Universal Robots URScript: MAIN_1.script

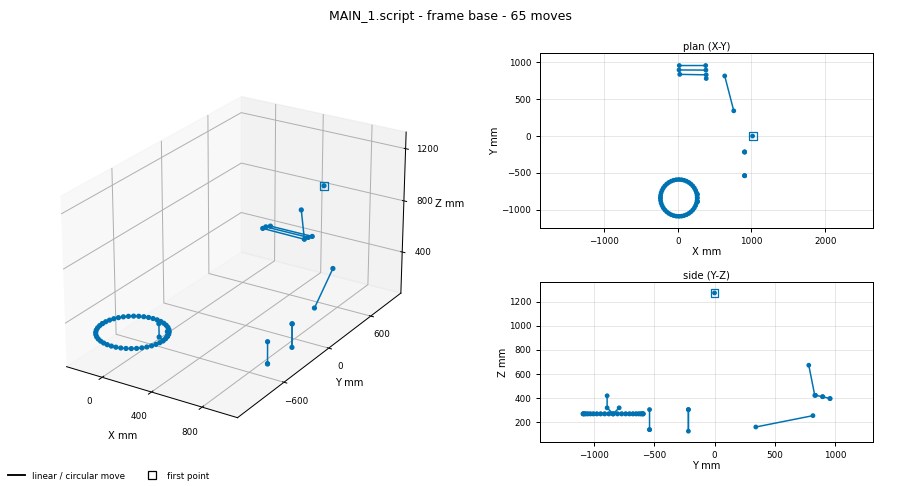
[picture p0: tool path of MAIN_1.script in frame base, 65 of 76 moves have a stored position in this frame; points joined in program order, loops and branches not executed]
def MAIN_1():
  # Global parameters:
  global speed_ms    = 0.300
  global speed_rads  = 0.750
  global accel_mss   = 3.000
  global accel_radss = 1.200
  global blend_radius_m = 0.001

  #--------------------------
  # Add any default subprograms here
  # For example, to drive a gripper as a program call:
  # def Gripper_Open():
  #   ...
  # end
  #
  # Example to drive a spray gun:
  def SprayOn(value):
    # use the value as an output:
    DO_SPRAY = 5
    if value == 0:
      set_standard_digital_out(DO_SPRAY, False)
    else:
      set_standard_digital_out(DO_SPRAY, True)
    end
  end

  # Example to drive an extruder:
  def Extruder(value):
    # use the value as an output:
    if value < 0:
      # stop extruder
    else:
      # start extruder
    end
  end

  # Example to move an external axis
  def MoveAxis(value):
    # use the value as an output:
    DO_AXIS_1 = 1
    DI_AXIS_1 = 1
    if value <= 0:
      set_standard_digital_out(DO_AXIS_1, False)

      # Wait for digital input to change state
      #while (get_standard_digital_in(DI_AXIS_1) != False):
      #  sync()
      #end
    else:
      set_standard_digital_out(DO_AXIS_1, True)

      # Wait for digital input to change state
      #while (get_standard_digital_in(DI_AXIS_1) != True):
      #  sync()
      #end
    end
  end
  #--------------------------

  # Subprogram PROG1_withaverylongnameandspecialcharacters
  def PROG1_withaverylongnameandspecialcharacters():
    # This is a subprogram call to PROG_1
    # set_reference(p[0.000000, 1.000000, 0.000000, 0.000000, 0.000000, 0.000000])
    set_tcp(p[0.000000, 0.000000, 0.200000, 0.000000, 0.000000, 0.000000])
    movej([-0.000000, 0.000000, 0.000000, 0.000000, 0.000000, -0.000000],accel_radss,speed_rads,0,blend_radius_m)
  end


  # Main program:
  # Program generated by RoboDK v5.6.9 for RoboDK Industrial on 26/02/2024 09:58:20
  # Using nominal kinematics.
  movej([-0.000000, 0.000000, 0.000000, 0.000000, 0.000000, -0.000000],accel_radss,speed_rads,0,0)
  movej([0.000000, 0.056047, -0.269194, 0.000000, 0.213148, -0.000000],accel_radss,speed_rads,0,0)
  movel(p[1.015000, 0.000000, 1.272000, 0.000000, 1.570796, 0.000000],accel_mss,speed_ms,0,blend_radius_m)
  set_standard_digital_out(5, True)
  set_standard_digital_out(5, True)
  set_standard_digital_out(5, 0.5)
  set_standard_digital_out(5, true)
  set_standard_digital_out(5, True)
  set_standard_digital_out(5, True)
  set_standard_digital_out(5, 0.5)
  set_standard_digital_out(5, true)
  var = val
  var = val
  while (get_standard_digital_in(5) != True):
    sync()
  end
  while (get_standard_digital_in(5) != True):
    sync()
  end
  while (get_standard_digital_in(5) != 0.5):
    sync()
  end
  while (get_standard_digital_in(5) != true):
    sync()
  end
  while (get_standard_digital_in(5) != True):
    sync()
  end
  while (var != val):
    sync()
  end
  while (var != val):
    sync()
  end
  popup("Message","Message",False,False,blocking=True)
  REMOTE_PROG_CALL_171()
  # CODE_INSERT_172
  # Insert Comment
  # set_reference(p[0.719013, -0.664003, 0.000000, 0.000000, 0.000000, 0.000000])
  set_tcp(p[0.129073, 0.000000, 0.085477, 0.000000, 0.398790, 0.000000])
  accel_radss = 13.963
  speed_rads  = 8.727
  blend_radius_m = 0.010
  movej([-0.511943, 0.814667, -0.000428, 0.463308, 0.443239, -0.901183],accel_radss,speed_rads,0,blend_radius_m)
  blend_radius_m = 0.000
  accel_mss   = 0.200
  speed_ms    = 0.100
  movel(p[0.906799, -0.538504, 0.139112, -0.000082, 3.138451, 0.000110],accel_mss,speed_ms,0,blend_radius_m)
  set_standard_digital_out(5, True)
  PICK_PART_111()
  blend_radius_m = 0.010
  accel_mss   = 0.600
  speed_ms    = 0.300
  movel([-0.511943, 0.814667, -0.000427, 0.463312, 0.443239, -0.901187],accel_mss,speed_ms,0,0)
  movel(p[0.906285, -0.216481, 0.305347, 0.000027, 3.138364, -0.000055],accel_mss,speed_ms,0,blend_radius_m)
  blend_radius_m = 0.000
  accel_mss   = 0.200
  speed_ms    = 0.100
  # MoveSearch command not implemented
  movel(p[0.906864, -0.216486, 0.126235, 0.000027, 3.138364, -0.000055],accel_mss,speed_ms,0,blend_radius_m)
  set_standard_digital_out(5, False)
  PLACE_PART_112()
  blend_radius_m = 0.010
  movel(p[0.906285, -0.216481, 0.305347, 0.000027, 3.138364, -0.000055],accel_mss,speed_ms,0,blend_radius_m)
  # set_reference(p[0.577670, 0.392250, 0.000000, 0.000000, 0.000000, 0.679972])
  blend_radius_m = 0.025
  accel_radss = 13.963
  speed_rads  = 8.727
  accel_mss   = 0.200
  speed_ms    = 0.100
  movej([0.910818, 0.797193, 0.120777, 1.164732, 0.347884, -1.618444],accel_radss,speed_rads,0,blend_radius_m)
  movec(p[0.884547, 0.696689, 0.231503, -2.018719, 2.221778, 0.218496],p[0.759304, 0.342075, 0.161073, -2.018719, 2.221778, 0.218496],accel_mss,speed_ms,blend_radius_m)
  # Circular movement using joint targets is not supported. Change the target type to cartesian or use a joint movement.
  blend_radius_m = 0.000
  accel_mss   = 0.200
  speed_ms    = 0.100
  movel(p[0.636704, 0.815780, 0.255156, -2.018719, 2.221778, 0.218496],accel_mss,speed_ms,0,blend_radius_m)
  movej([-0.000000, 0.000000, 0.000000, 0.000000, 0.000000, -0.000000],accel_radss,speed_rads,0,0)
  # set_reference(p[0.000000, 0.782714, 0.377610, 0.000000, 0.000000, 0.000000])
  movej([1.547688, 0.516645, -0.112204, -0.034631, 0.863575, 0.079372],accel_radss,speed_rads,0,0)
  movel(p[0.019898, 0.957021, 0.396618, 2.079600, -2.265750, 0.107759],accel_mss,speed_ms,0,blend_radius_m)
  movel(p[0.378402, 0.957130, 0.396607, 2.079600, -2.265750, 0.107759],accel_mss,speed_ms,0,blend_radius_m)
  movel(p[0.380996, 0.895077, 0.412492, 1.963520, -2.143933, 0.343573],accel_mss,speed_ms,0,blend_radius_m)
  movel(p[0.016551, 0.897073, 0.411836, 1.963520, -2.143933, 0.343573],accel_mss,speed_ms,0,blend_radius_m)
  movel(p[0.026434, 0.837238, 0.423682, -2.078092, 2.285598, 0.087159],accel_mss,speed_ms,0,blend_radius_m)
  movel(p[0.385448, 0.830764, 0.422747, -2.018705, 2.221797, 0.218488],accel_mss,speed_ms,0,blend_radius_m)
  movel(p[0.385448, 0.781089, 0.672861, -2.018705, 2.221797, 0.218488],accel_mss,speed_ms,0,blend_radius_m)
  movej([-0.000000, 0.000000, 0.000000, 0.000000, 0.000000, -0.000000],accel_radss,speed_rads,0,0)
  EVENT_PROG_START_101()
  blend_radius_m = 0.001
  speed_ms    = 1.000
  # set_reference(p[0.013637, -0.840080, 0.000000, 0.000000, 0.000000, -1.570796])
  # Show Tool 1
  movej([-1.188400, 0.422403, 0.467495, 0.666950, 0.631839, -1.724322],accel_radss,speed_rads,0,0)
  EVENT_PATH_APPROACH_102()
  movel(p[0.266896, -0.790185, 0.319999, 0.000002, 3.135432, -0.000684],accel_mss,speed_ms,0,blend_radius_m)
  movel(p[0.263637, -0.840080, 0.270000, 0.000002, 3.135432, -0.000684],accel_mss,speed_ms,0,blend_radius_m)
  EVENT_PATH_START_103()
  speed_ms    = 0.050
  movel(p[0.261092, -0.875659, 0.270000, 0.000006, 3.135571, -0.002052],accel_mss,speed_ms,0,blend_radius_m)
  movel(p[0.253510, -0.910513, 0.270000, -0.000018, 3.135814, -0.003393],accel_mss,speed_ms,0,blend_radius_m)
  movel(p[0.241045, -0.943934, 0.270000, -0.000015, 3.136179, -0.004625],accel_mss,speed_ms,0,blend_radius_m)
  movel(p[0.223950, -0.975240, 0.270000, -0.000013, 3.136648, -0.005803],accel_mss,speed_ms,0,blend_radius_m)
  movel(p[0.202574, -1.003795, 0.270000, -0.000012, 3.137222, -0.006844],accel_mss,speed_ms,0,blend_radius_m)
  movel(p[0.177352, -1.029017, 0.270000, -0.000013, 3.137883, -0.007749],accel_mss,speed_ms,0,blend_radius_m)
  movel(p[0.148797, -1.050393, 0.270000, -0.000015, 3.138614, -0.008518],accel_mss,speed_ms,0,blend_radius_m)
  movel(p[0.117491, -1.067488, 0.270000, -0.000018, 3.139415, -0.009096],accel_mss,speed_ms,0,blend_radius_m)
  movel(p[0.084070, -1.079953, 0.270000, 0.000006, 3.140269, -0.009482],accel_mss,speed_ms,0,blend_radius_m)
  movel(p[0.049216, -1.087535, 0.270000, 0.000002, 3.141141, -0.009676],accel_mss,speed_ms,0,blend_radius_m)
  movel(p[0.013637, -1.090080, 0.270000, 0.000002, -3.141141, 0.009676],accel_mss,speed_ms,0,blend_radius_m)
  movel(p[-0.021942, -1.087535, 0.270000, 0.000006, -3.140269, 0.009482],accel_mss,speed_ms,0,blend_radius_m)
  movel(p[-0.056796, -1.079953, 0.270000, -0.000018, -3.139415, 0.009096],accel_mss,speed_ms,0,blend_radius_m)
  movel(p[-0.090217, -1.067488, 0.270000, -0.000015, -3.138614, 0.008518],accel_mss,speed_ms,0,blend_radius_m)
  movel(p[-0.121523, -1.050393, 0.270000, -0.000013, -3.137883, 0.007749],accel_mss,speed_ms,0,blend_radius_m)
  movel(p[-0.150078, -1.029017, 0.270000, -0.000012, -3.137222, 0.006844],accel_mss,speed_ms,0,blend_radius_m)
  movel(p[-0.175300, -1.003795, 0.270000, -0.000013, -3.136648, 0.005803],accel_mss,speed_ms,0,blend_radius_m)
  movel(p[-0.196676, -0.975240, 0.270000, -0.000015, -3.136161, 0.004653],accel_mss,speed_ms,0,blend_radius_m)
  movel(p[-0.213771, -0.943934, 0.270000, -0.000018, -3.135796, 0.003393],accel_mss,speed_ms,0,blend_radius_m)
  movel(p[-0.226236, -0.910513, 0.270000, 0.000006, -3.135553, 0.002052],accel_mss,speed_ms,0,blend_radius_m)
  movel(p[-0.233818, -0.875659, 0.270000, 0.000002, -3.135432, 0.000684],accel_mss,speed_ms,0,blend_radius_m)
  movel(p[-0.236363, -0.840080, 0.270000, 0.000002, -3.135432, 0.000684],accel_mss,speed_ms,0,blend_radius_m)
  movel(p[-0.236363, -0.840080, 0.270000, -0.000002, -3.135432, -0.000684],accel_mss,speed_ms,0,0.000)
  movel(p[-0.233818, -0.804501, 0.270000, -0.000006, -3.135553, -0.002052],accel_mss,speed_ms,0,blend_radius_m)
  movel(p[-0.226236, -0.769647, 0.270000, 0.000018, -3.135814, -0.003393],accel_mss,speed_ms,0,blend_radius_m)
  movel(p[-0.213771, -0.736226, 0.270000, 0.000015, -3.136179, -0.004625],accel_mss,speed_ms,0,blend_radius_m)
  movel(p[-0.196676, -0.704920, 0.270000, 0.000013, -3.136648, -0.005803],accel_mss,speed_ms,0,blend_radius_m)
  movel(p[-0.175300, -0.676365, 0.270000, 0.000012, -3.137222, -0.006844],accel_mss,speed_ms,0,blend_radius_m)
  movel(p[-0.150078, -0.651143, 0.270000, 0.000013, -3.137883, -0.007749],accel_mss,speed_ms,0,blend_radius_m)
  movel(p[-0.121523, -0.629767, 0.270000, 0.000015, -3.138632, -0.008491],accel_mss,speed_ms,0,blend_radius_m)
  movel(p[-0.090217, -0.612672, 0.270000, 0.000018, -3.139433, -0.009068],accel_mss,speed_ms,0,blend_radius_m)
  movel(p[-0.056796, -0.600207, 0.270000, -0.000006, -3.140269, -0.009482],accel_mss,speed_ms,0,blend_radius_m)
  movel(p[-0.021942, -0.592625, 0.270000, -0.000002, -3.141141, -0.009676],accel_mss,speed_ms,0,blend_radius_m)
  movel(p[0.013637, -0.590080, 0.270000, -0.000002, 3.141141, 0.009676],accel_mss,speed_ms,0,blend_radius_m)
  movel(p[0.049216, -0.592625, 0.270000, -0.000006, 3.140269, 0.009454],accel_mss,speed_ms,0,blend_radius_m)
  movel(p[0.084070, -0.600207, 0.270000, 0.000018, 3.139433, 0.009068],accel_mss,speed_ms,0,blend_radius_m)
  movel(p[0.117491, -0.612672, 0.270000, 0.000015, 3.138614, 0.008518],accel_mss,speed_ms,0,blend_radius_m)
  movel(p[0.148797, -0.629767, 0.270000, 0.000013, 3.137883, 0.007749],accel_mss,speed_ms,0,blend_radius_m)
  movel(p[0.177352, -0.651143, 0.270000, 0.000012, 3.137222, 0.006844],accel_mss,speed_ms,0,blend_radius_m)
  movel(p[0.202574, -0.676365, 0.270000, 0.000013, 3.136648, 0.005803],accel_mss,speed_ms,0,blend_radius_m)
  movel(p[0.223950, -0.704920, 0.270000, 0.000015, 3.136179, 0.004625],accel_mss,speed_ms,0,blend_radius_m)
  movel(p[0.241045, -0.736226, 0.270000, 0.000018, 3.135796, 0.003393],accel_mss,speed_ms,0,blend_radius_m)
  movel(p[0.253510, -0.769647, 0.270000, -0.000006, 3.135553, 0.002052],accel_mss,speed_ms,0,blend_radius_m)
  movel(p[0.261092, -0.804501, 0.270000, -0.000002, 3.135432, 0.000684],accel_mss,speed_ms,0,blend_radius_m)
  movel(p[0.263637, -0.840080, 0.270000, -0.000002, 3.135432, 0.000684],accel_mss,speed_ms,0,blend_radius_m)
  speed_ms    = 1.000
  EVENT_PATH_FINISH_105()
  movel(p[0.266895, -0.889975, 0.319999, -0.000002, 3.135432, 0.000684],accel_mss,speed_ms,0,blend_radius_m)
  movel(p[0.266279, -0.890019, 0.419997, -0.000002, 3.135432, 0.000684],accel_mss,speed_ms,0,blend_radius_m)
  EVENT_PATH_RETRACT_106()
  EVENT_PROG_FINISH_107()
  # set_reference(p[0.719013, -0.664003, 0.000000, 0.000000, 0.000000, 0.000000])
  movej([-0.511943, 0.814667, -0.000428, 0.463308, 0.443239, -0.901183],accel_radss,speed_rads,0,blend_radius_m)
  sleep(1.250)
  movel(p[0.906799, -0.538504, 0.139112, -0.000082, 3.138451, 0.000110],accel_mss,speed_ms,0,blend_radius_m)
  while (get_standard_digital_in(1) != True):
    sync()
  end
  movel(p[0.906277, -0.538516, 0.305356, 0.000000, 3.138381, -0.000000],accel_mss,speed_ms,0,blend_radius_m)
  PROG1_withaverylongnameandspecialcharacters()
  # End of main program
end

MAIN_1()
